Staubli VAL3: changeBckColorLabel.pgx

public program changeBckColorLabel(utLabel x_uUtLabel, string x_sColor)
begin
  // change the BackGround color -> using userPageSet
  userPageSet(x_uUtLabel.Common.sPage,x_uUtLabel.Common.sID,"style.backgroundColor",x_sColor)
end
